Staubli VAL3: refreshlist.pgx

program refreshlist()
  local num l_nSize
  local string l_sTrajList
  local num l_i
  local num l_nCount
begin
  call trajectory:getTrajSize(l_nSize)
  call trajectory:getTrajList(sTrajList)
  //page
  if l_nSize<50
    nPageNum=1
  else
    nPageNum=roundUp(l_nSize/49)
  endIf

  //list
  if nPageNum==1
    if l_nSize<1
      for l_i = 0 to size(sList)-1
        sList[l_i]=""
      endFor
    else
      resize(sList,1,l_nSize)
      for l_i = 0 to size(sList)-1
        sList[l_i]=""
      endFor
      for l_i = 0 to l_nSize-1
        sList[l_i]=sTrajList[l_i]
      endFor
    endIf

  else
    if nPageIndex<nPageNum-1
      resize(sList,1,49)
      for l_i = 0 to size(sList)-1
        sList[l_i]=sTrajList[nPageIndex*49+l_i]
      endFor
    else
      for l_i = 0 to size(sList)-1
        sList[l_i]=""
      endFor
      if l_nSize%49==0
        l_nCount=49
      else
        l_nCount=l_nSize%49
      endIf
      resize(sList,1,l_nCount)
      for l_i = 0 to l_nCount-1
        sList[l_i]=sTrajList[l_i+nPageIndex*49]
      endFor
    endIf
  endIf
  userPageBind("traj","lst1","options",sList,size(sList),"r")
  sPageIndex=toString("",nPageIndex+1)
  sPageNum=toString("",nPageNum)
end
